// TIA Portal V21 export
FUNCTION_BLOCK "HMI_Bedienung_Animationen"   // FB3, FBD
{ S7_Optimized_Access := 'TRUE' }
// Dieser Baustein ist nur für die Bedienbarkeit der HMI zuständig. Um eine Funktion (z.B. Jog-Mode) auf der HMI zu aktivieren, müssen Bedigungen erfüllt sein.
// stored: MemoryReserve 100, SetENOAutomatically false
   VAR
      "ActVel_h_%" : LReal;
      "ActVel_v_%" : LReal;
   END_VAR
BEGIN

REGION Network 1: einschubachse eingefahren
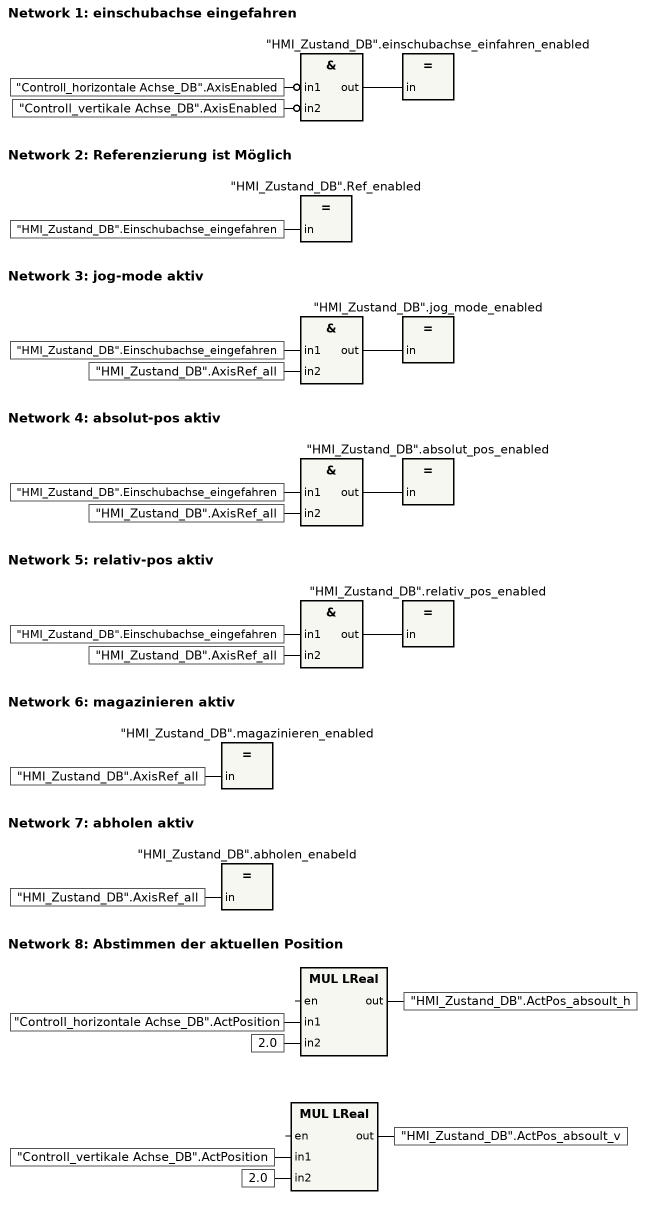
   "HMI_Zustand_DB".einschubachse_einfahren_enabled := NOT "Controll_horizontale Achse_DB".AxisEnabled AND NOT "Controll_vertikale Achse_DB".AxisEnabled;
END_REGION

REGION Network 2: Referenzierung ist Möglich
   "HMI_Zustand_DB".Ref_enabled := "HMI_Zustand_DB".Einschubachse_eingefahren;
END_REGION

REGION Network 3: jog-mode aktiv
   "HMI_Zustand_DB".jog_mode_enabled := "HMI_Zustand_DB".Einschubachse_eingefahren AND "HMI_Zustand_DB".AxisRef_all;
END_REGION

REGION Network 4: absolut-pos aktiv
   "HMI_Zustand_DB".absolut_pos_enabled := "HMI_Zustand_DB".Einschubachse_eingefahren AND "HMI_Zustand_DB".AxisRef_all;
END_REGION

REGION Network 5: relativ-pos aktiv
   "HMI_Zustand_DB".relativ_pos_enabled := "HMI_Zustand_DB".Einschubachse_eingefahren AND "HMI_Zustand_DB".AxisRef_all;
END_REGION

REGION Network 6: magazinieren aktiv
   "HMI_Zustand_DB".magazinieren_enabled := "HMI_Zustand_DB".AxisRef_all;
END_REGION

REGION Network 7: abholen aktiv
   "HMI_Zustand_DB".abholen_enabeld := "HMI_Zustand_DB".AxisRef_all;
END_REGION

REGION Network 8: Abstimmen der aktuellen Position
   // Die Aktuelle Psoition wird hier bearbeitet so das Anzeige und HRL ident sind.
   "HMI_Zustand_DB".ActPos_absoult_h := "Controll_horizontale Achse_DB".ActPosition * 2.0;
   "HMI_Zustand_DB".ActPos_absoult_v := "Controll_vertikale Achse_DB".ActPosition * 2.0;
END_REGION

REGION Network 9: Berechnung der Animationswerte für horizontale Achse
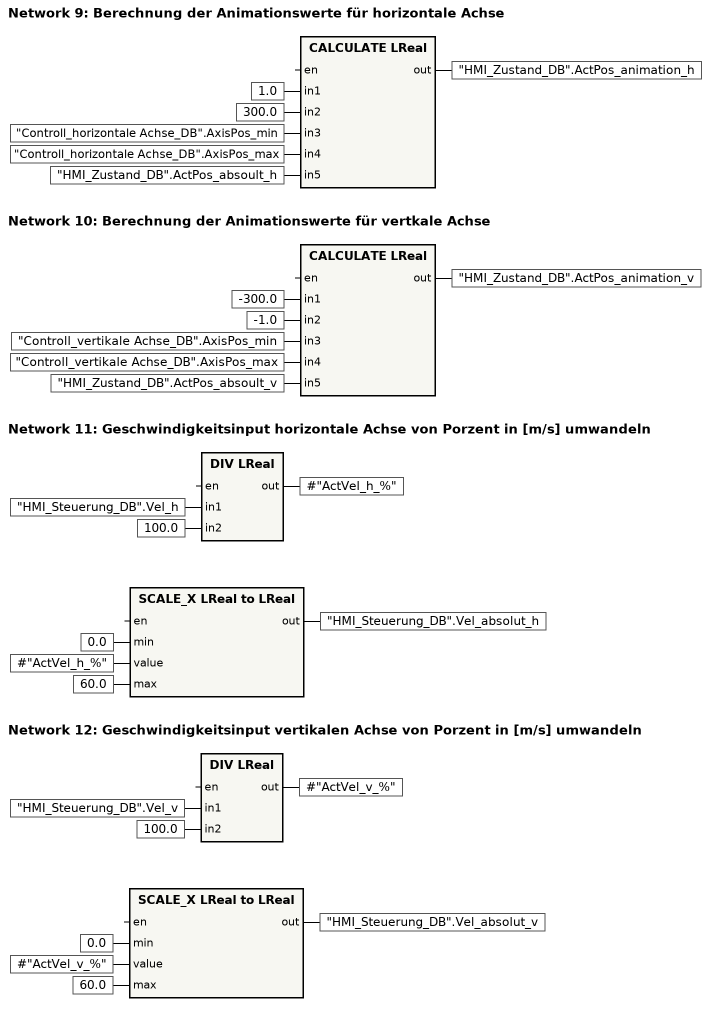
   "HMI_Zustand_DB".ActPos_animation_h := (1.0-(("Controll_horizontale Achse_DB".AxisPos_max-"HMI_Zustand_DB".ActPos_absoult_h)/("Controll_horizontale Achse_DB".AxisPos_max+ABS("Controll_horizontale Achse_DB".AxisPos_min))))*300.0;
END_REGION

REGION Network 10: Berechnung der Animationswerte für vertkale Achse
   "HMI_Zustand_DB".ActPos_animation_v := (-"HMI_Zustand_DB".ActPos_absoult_v/("Controll_vertikale Achse_DB".AxisPos_max-"Controll_vertikale Achse_DB".AxisPos_min))*((-1.0)-(-300.0));
END_REGION

REGION Network 11: Geschwindigkeitsinput horizontale Achse von Porzent in [m/s] umwandeln
   #"ActVel_h_%" := "HMI_Steuerung_DB".Vel_h / 100.0;
   "HMI_Steuerung_DB".Vel_absolut_h := SCALE_X(MIN := 0.0, VALUE := #"ActVel_h_%", MAX := 60.0);
END_REGION

REGION Network 12: Geschwindigkeitsinput vertikalen Achse von Porzent in [m/s] umwandeln
   #"ActVel_v_%" := "HMI_Steuerung_DB".Vel_v / 100.0;
   "HMI_Steuerung_DB".Vel_absolut_v := SCALE_X(MIN := 0.0, VALUE := #"ActVel_v_%", MAX := 60.0);
END_REGION
END_FUNCTION_BLOCK
